// TIA Portal V21 export
// export: Created 2026-10-12T11:32:11.3403395Z, ExportSetting WithDefaults, DisplayName Totally Integrated Automation Portal, DisplayVersion V21, DisplayName STEP 7 Professional, DisplayVersion V21, DisplayName STEP 7 Safety, DisplayVersion V21, DisplayName Tech WebApplication, DisplayVersion V21, DisplayName WinCC Basic/Comfort/Advanced, DisplayVersion V21, DisplayName WinCC Unified, DisplayVersion V21
ORGANIZATION_BLOCK "Main"   // OB1, LAD, ProgramCycle
TITLE = "Main Program Sweep (Cycle)"
{ S7_Optimized_Access := 'TRUE' }
VERSION : 0.1
// stored: AutoNumber true, IsIECCheckEnabled false, SetENOAutomatically false
   VAR_INPUT
      Initial_Call : Bool;   // Initial call of this OB
      Remanence : Bool;   // =True, if remanent data are available
   END_VAR
BEGIN

REGION Network 1
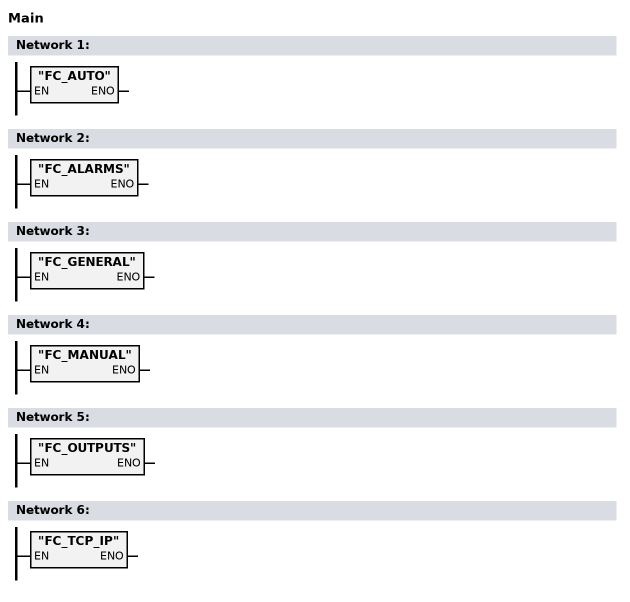
   RUNG wire#powerrail
      "FC_AUTO"()
   END_RUNG
   // the same network as SCL:
   "FC_AUTO"();
END_REGION

REGION Network 2
   RUNG wire#powerrail
      "FC_ALARMS"()
   END_RUNG
   // the same network as SCL:
   "FC_ALARMS"();
END_REGION

REGION Network 3
   RUNG wire#powerrail
      "FC_GENERAL"()
   END_RUNG
   // the same network as SCL:
   "FC_GENERAL"();
END_REGION

REGION Network 4
   RUNG wire#powerrail
      "FC_MANUAL"()
   END_RUNG
   // the same network as SCL:
   "FC_MANUAL"();
END_REGION

REGION Network 5
   RUNG wire#powerrail
      "FC_OUTPUTS"()
   END_RUNG
   // the same network as SCL:
   "FC_OUTPUTS"();
END_REGION

REGION Network 6
   RUNG wire#powerrail
      "FC_TCP_IP"()
   END_RUNG
   // the same network as SCL:
   "FC_TCP_IP"();
END_REGION
END_ORGANIZATION_BLOCK
